{region 'Documentation'}
(*!
<summary>Rejects a missing Start reaction at the first-slot boundary without starting the next slot.</summary>
<description>
Child 1 completes immediately. Child 2 is then admitted but remains Idle.
The pending Start must be rejected once, its reservation released and child 3 left
untouched in slot 2. Repeated calls must preserve the Error without repeating diagnostics.
</description>
*)
{endregion}
FUNCTION_BLOCK Test_SlotsMissingStartReaction EXTENDS OrchestrationTestBase

SUPER^();

{region 'Documentation'}
(*!
<summary>Defines boundary stimuli and expected child requests, reservation cleanup and isolated diagnostics.</summary>
*)
{endregion}
METHOD PROTECTED ConfigureScenario
FChildSlots[1] := 1;
FChildSlots[2] := 1;
FChildSlots[3] := 2;
FStepCount := 5;

{region "01 - Observe initial readiness"}
FSteps[1].Task := E_OrchestratorTask.Idle;
FSteps[1].ExpectedReady := TRUE;
FSteps[1].MaxActiveChildCount := 0;
{endregion}

{region "02 - Child 1 completes immediately after Start"}
FSteps[2].Children[1].State := E_State.Completed;
FSteps[2].Children[1].Ready := FALSE;
FSteps[2].Children[1].Complete := TRUE;
FSteps[2].Children[1].Result := E_Result.Passed;
FSteps[2].ExpectedStartChild := 1;
FSteps[2].ExpectedSlot := 1;
FSteps[2].ExpectedReservations[1] := 1;
FSteps[2].MaxActiveChildCount := 1;
{endregion}

{region "03 - Start child 2 but retain its Idle observation"}
FSteps[3].Children[1].State := E_State.Completed;
FSteps[3].Children[1].Ready := FALSE;
FSteps[3].Children[1].Complete := TRUE;
FSteps[3].Children[1].Result := E_Result.Passed;
FSteps[3].ExpectedStartChild := 2;
FSteps[3].ExpectedSlot := 1;
FSteps[3].ExpectedReservations[2] := 1;
FSteps[3].ExpectedReleasedEntries[1] := 1;
FSteps[3].MaxActiveChildCount := 1;
{endregion}

{region "04 - Reject the missing reaction and release the pending reservation"}
FSteps[4].Children[1].State := E_State.Completed;
FSteps[4].Children[1].Ready := FALSE;
FSteps[4].Children[1].Complete := TRUE;
FSteps[4].Children[1].Result := E_Result.Passed;
FSteps[4].ExpectedSlot := 1;
FSteps[4].ExpectedResult := E_Result.Error;
FSteps[4].ExpectedDiagnosticCount := 1;
FSteps[4].ExpectedReleasedEntries[2] := 1;
FSteps[4].MaxActiveChildCount := 0;
{endregion}

{region "05 - Keep the next slot blocked without repeating the diagnostic"}
FSteps[5].Children[1].State := E_State.Completed;
FSteps[5].Children[1].Ready := FALSE;
FSteps[5].Children[1].Complete := TRUE;
FSteps[5].Children[1].Result := E_Result.Passed;
FSteps[5].ExpectedSlot := 1;
FSteps[5].ExpectedResult := E_Result.Error;
FSteps[5].ExpectedDiagnosticCount := 1;
FSteps[5].MaxActiveChildCount := 0;
{endregion}
END_METHOD

END_FUNCTION_BLOCK

(* stored: Version 1.1.0.1
   POU Test_SlotsMissingStartReaction: Id {4d7a55d0-f7ab-4b0e-9148-1f1a5418fd31}, SpecialFunc None
   Folder Internal: Id {adcb4610-53ab-4cfa-8e99-000000000004}
   Method ConfigureScenario: Id {adcb4620-53ab-4cfa-8e99-000000000004} *)
